// TIA Portal V20 export
Screen "Pop-up_StyleConfigLocal"  653x462
